(* IEC 61131-3 sources: plc-vscode/tests/st/test-ready/rusty/tests/lit/correctness/functions, 6 files *)

(* ---- sizeof_test.st ---- *)
// RUN: (%COMPILE %s && %RUN) | %CHECK %s

CLASS MyClass
    VAR
    x, y: INT; // 4 bytes
    END_VAR
END_CLASS

TYPE MyStruct: STRUCT
    a: BYTE; // 8bit - offset 0 -> 1 byte
    b: DWORD; // 32bit - offset 32 -> 8 bytes
    c: WORD; // 16bit - offset 64 -> 10 bytes
    d: LWORD; // 64bit - offset 128 -> 24 bytes
END_STRUCT END_TYPE

FUNCTION main
    VAR
        s1: SINT;
        s2: INT;
        s3: DINT;
        s4: LINT;
        s5: USINT;
        s6: UDINT;
        s7: ULINT;
        s8: LINT;
    END_VAR

    VAR_TEMP
        t1: MyStruct;
        t2: STRING;
        t3: WCHAR;
        t4: MyClass;
        t5: LREAL;
        t6: BOOL;
    END_VAR

    s1 := SIZEOF(t6);
    s2 := SIZEOF(s2);
    s3 := SIZEOF(t5);
    s4 := SIZEOF(t1);
    s5 := SIZEOF(REF(s1));
    s6 := SIZEOF(t2);
    s7 := SIZEOF(t3);
    s8 := SIZEOF(t4);

    printf('s1 = %d$N', s1); // CHECK: s1 = 1
    printf('s2 = %d$N', s2); // CHECK: s2 = 2
    printf('s3 = %d$N', s3); // CHECK: s3 = 8
    printf('s4 = %d$N', s4); // CHECK: s4 = 24
    printf('s5 = %d$N', s5); // CHECK: s5 = 8
    printf('s6 = %d$N', s6); // CHECK: s6 = 81
    printf('s7 = %d$N', s7); // CHECK: s7 = 2
    printf('s8 = %d$N', s8); // CHECK: s8 = 16
END_FUNCTION

(* ---- mixed_implicit_explicit_trailing_defaults.st ---- *)
// RUN: (%COMPILE %s && %RUN) | %CHECK %s

// Runtime check that trailing defaults fill correctly when combined with mixed
// positional/named args. The resolver's "skip named slots" rule for positionals
// must leave genuinely-omitted trailing slots to pick up the declared default.
//
// Related gap pinned in `mixed_implicit_explicit_non_trailing_default_is_rejected`:
// non-trailing defaults (e.g. `a, b := 1, c`) are NOT accepted. IEC 61131-3
// semantics would suggest they should, but RuSTy rejects them today.

FUNCTION myfunc : DINT
VAR_INPUT
    a : DINT;
    b : DINT := 1000;
    c : DINT := 100;
END_VAR
    myfunc := a * 10000 + b * 10 + c;
END_FUNCTION

FUNCTION main
VAR
    r1, r2, r3, r4 : DINT;
END_VAR
    // one positional, rest defaulted
    r1 := myfunc(5);                 // a=5  b=1000 c=100 -> 60100

    // positional + named, c defaulted
    r2 := myfunc(5, b := 2);         // a=5  b=2    c=100 -> 50120

    // named + positional, c defaulted (positional 2 fills b via skip-named-slots)
    r3 := myfunc(a := 5, 2);         // a=5  b=2    c=100 -> 50120

    // all supplied, defaults overridden
    r4 := myfunc(5, 2, 3);           // a=5  b=2    c=3   -> 50023

    printf('r1=%d$N', r1); // CHECK: r1=60100
    printf('r2=%d$N', r2); // CHECK: r2=50120
    printf('r3=%d$N', r3); // CHECK: r3=50120
    printf('r4=%d$N', r4); // CHECK: r4=50023
END_FUNCTION

(* ---- direct_call_on_function_block_array_access.st ---- *)
// RUN: (%COMPILE %s && %RUN) | %CHECK %s

FUNCTION_BLOCK foo
    VAR_INPUT
        i: INT;
    END_VAR
    VAR
        x: INT;
    END_VAR

    x := i;
END_FUNCTION_BLOCK

FUNCTION main
    VAR
        f: ARRAY[1..2] OF foo;
        x: INT;
        y: INT;
    END_VAR

    f[1](i := 10);
    x := f[1].x;

    f[2](i := 20);
    y := f[2].x;

    printf('x = %d$N', x); // CHECK: x = 10
    printf('y = %d$N', y); // CHECK: y = 20
END_FUNCTION

(* ---- function_block_instances_save_state_per_instance.st ---- *)
// RUN: (%COMPILE %s && %RUN) | %CHECK %s

FUNCTION_BLOCK foo
    VAR_INPUT
        i: INT;
    END_VAR

    i := i + 1;
END_FUNCTION_BLOCK

FUNCTION main
    VAR
        f: foo;
        j: foo;
    END_VAR

    f();
    f();
    j(4);
    j();
    j();

    printf('f.i = %d$N', f.i); // CHECK: f.i = 2
    printf('j.i = %d$N', j.i); // CHECK: j.i = 7
END_FUNCTION

(* ---- function_block_instances_save_state_per_instance_2.st ---- *)
// RUN: (%COMPILE %s && %RUN) | %CHECK %s
FUNCTION_BLOCK Baz
    VAR_INPUT
        i: INT;
    END_VAR

    i := i + 1;
END_FUNCTION_BLOCK

FUNCTION_BLOCK foo
    VAR_INPUT
        i: INT;
        baz: Baz;
    END_VAR
END_FUNCTION_BLOCK

FUNCTION main
    VAR
        f: foo;
        j: foo;
    END_VAR

    f.baz.i := f.baz.i + 1;
    f.baz.i := f.baz.i + 1;

    j.baz.i := j.baz.i + 1;
    j.baz.i := j.baz.i + 1;
    j.baz.i := j.baz.i + 1;
    j.baz.i := j.baz.i + 1;

    printf('f.baz.i = %d$N', f.baz.i); // CHECK: f.baz.i = 2
    printf('j.baz.i = %d$N', j.baz.i); // CHECK: j.baz.i = 4
END_FUNCTION

(* ---- mixed_implicit_explicit_args.st ---- *)
// RUN: (%COMPILE %s && %RUN) | %CHECK %s

// Verify that mixing positional and named arguments compiles and produces
// correct results at runtime.

FUNCTION add3 : INT
VAR_INPUT
    a : INT;
    b : INT;
    c : INT;
END_VAR
    add3 := a * 100 + b * 10 + c;
END_FUNCTION

FUNCTION_BLOCK Counter
VAR_INPUT
    step  : INT;
    start : INT;
END_VAR
VAR_OUTPUT
    val : INT;
END_VAR
    val := start + step;
END_FUNCTION_BLOCK

FUNCTION main
VAR
    r1, r2, r3, r4, r5 : INT;
    fb : Counter;
END_VAR
    // positional before named
    r1 := add3(1, b := 20, c := 3);   // a=1  b=20 c=3  -> 123  wait, 1*100+20*10+3 = 303
    // named before positional
    r2 := add3(a := 10, 2, c := 3);   // a=10 b=2  c=3  -> 1023
    // named non-first param, rest positional
    r3 := add3(b := 20, 1, 3);        // a=1  b=20 c=3  -> 303
    // only one named, two positional
    r4 := add3(10, 2, c := 30);       // a=10 b=2  c=30 -> 1050
    // function block: positional input + named output
    fb(1, start := 10, val => r5);    // step=1 start=10 -> val=11

    printf('r1=%d$N', r1); // CHECK: r1=303
    printf('r2=%d$N', r2); // CHECK: r2=1023
    printf('r3=%d$N', r3); // CHECK: r3=303
    printf('r4=%d$N', r4); // CHECK: r4=1050
    printf('r5=%d$N', r5); // CHECK: r5=11
END_FUNCTION
